    rq_activate_all_grippers(True)
    # end: URCap Program Node
  end
  $ 60 "zero_ftsensor()"
  zero_ftsensor()
  $ 61 "EXTT"
  $ 62 "Set GRP_3F_Enable=Off"
  set_standard_digital_out(4, False)
  $ 63 "Set BarcodeTrigger=Off"
  set_standard_digital_out(6, False)
  $ 64 "Set GRP_3F_Decap=Off"
  set_standard_digital_out(3, False)
  $ 65 "Set GRP_3F_Cap=Off"
  set_standard_digital_out(2, False)
  $ 66 "Set GRP_3F_Open=Off"
  set_standard_digital_out(5, False)
  $ 67 "PSE_T≔get_tool_free_pose(dir=[0,0,0.150], move_in_base_frame=True)"
  global PSE_T=get_tool_free_pose(dir=[0,0,0.150], move_in_base_frame=True)
  $ 68 "If is_reachable(Base_const, [PSE_T])"
  if (is_reachable(p[0.0,0.0,0.0,0.0,0.0,0.0], [PSE_T])):
    $ 69 "MoveL"
    $ 70 "PSE_T" "breakAfter"
    movel(PSE_T, a=1.2, v=0.15)
  end
  $ 71 "powder dispensing variable init"
  $ 72 "Start_thread≔ False "
  global Start_thread=  False
  $ 73 "vib_thread≔ False "
  global vib_thread=  False
  $ 74 "kp≔0.0002"
  global kp=0.0002
  $ 75 "ki≔0.001"
  global ki=0.001
  $ 76 "kd≔0.01"
  global kd=0.01
  $ 77 "dt≔0.05"
  global dt=0.05
  $ 78 "Integral_error≔0"
  global Integral_error=0
  $ 79 "current_error≔0"
  global current_error=0
  $ 80 "previous_error≔0"
  global previous_error=0
  $ 81 "tilt_increment≔0"
  global tilt_increment=0
  $ 82 "tilt_angle≔-1"
  global tilt_angle=-1
  $ 83 "diff≔0"
  global diff=0
  $ 84 "current_pose≔get_actual_tcp_pose()"
  global current_pose= get_actual_tcp_pose ()
  while (True):
    $ 85 "Robot Program"
    $ 86 "MAIN"
    $ 87 "command_manager(external_control='uGO', cond_suspend=(ITM_Manipulated and AMR_AtTarget and AMR_Charging and AMR_Battery<40), cond_unsuspend=(AMR_Battery≟60))"
    command_manager(external_control="uGO", cond_suspend=(ITM_Manipulated  and  AMR_AtTarget  and  AMR_Charging  and  AMR_Battery<40), cond_unsuspend=(AMR_Battery == 60))
    $ 88 "log_state(STATE_Info)"
    log_state(STATE_Info)
    $ 89 "Switch STATE"
    switch_1 = STATE
    $ 90 "Case 1"
    if (1 == switch_1):
      $ 91 "Stopping"
      $ 92 "STATE_Info≔'Stopping'"
      global STATE_Info="Stopping"
      $ 93 "end_freedrive_mode()"
      end_freedrive_mode()
      $ 94 "Set"
      set_tcp(p[0.0,0.0,0.161,3.1415,0.0,0.0])
      $ 95 "PSE_T≔get_tool_free_pose(dir=[0,0,0.150], move_in_base_frame=True)"
      global PSE_T=get_tool_free_pose(dir=[0,0,0.150], move_in_base_frame=True)
      $ 96 "If is_reachable(Base_const, [PSE_T])"
      if (is_reachable(p[0.0,0.0,0.0,0.0,0.0,0.0], [PSE_T])):
        $ 97 "MoveL"
        $ 98 "PSE_T" "breakAfter"
        movel(PSE_T, a=1.2, v=0.15)
      end
      $ 99 "do_transition(keep_rxry=OBJ_Picked, r=0)"
      do_transition(keep_rxry=OBJ_Picked, r=0)
      $ 108 "Call Sub_AMR_MiR_V3"
      Sub_AMR_MiR_V3()
      $ 109 "If stopping() and AMR_Done"
      if (stopping()  and  AMR_Done):
        $ 110 "STATE≔2"
        global STATE=2
        $ 111 "ugo_update_outputs()"
        ugo_update_outputs()
      end
    elif (2 == switch_1):
      $ 112 "Case 2"
      $ 113 "Stopped"
      $ 114 "STATE_Info≔'Stopped'"
      global STATE_Info="Stopped"
      $ 115 "Call Sub_AMR_MiR_V3"
      Sub_AMR_MiR_V3()
      $ 116 "If CMD_Reset  or PB_Start"
      if (CMD_Reset   or  get_standard_digital_in(0)):
        $ 117 "STATE≔3"
        global STATE=3
        $ 118 "ugo_update_outputs()"
        ugo_update_outputs()
      end
    elif (3 == switch_1):
      $ 119 "Case 3"
      $ 120 " Resetting"
      $ 121 "STATE_Info≔'Resetting'"
      global STATE_Info="Resetting"
      $ 122 "uML"
      $ 123 "reset_error()"
      reset_error()
      $ 124 "reset_warning()"
      reset_warning()
      $ 125 "PROCESS_Step≔0"
      global PROCESS_Step=0
      $ 126 "PROCESS_Info≔''"
      global PROCESS_Info=""
      $ 127 "ARM_Referenced≔ False "
      global ARM_Referenced=  False
      $ 128 "WRK_Done≔ False "
      global WRK_Done=  False
      $ 129 "ITM_Prepared≔ False "
      global ITM_Prepared=  False
      $ 130 "ITM_Manipulated≔ False "
      global ITM_Manipulated=  False
      $ 131 "STP≔0"
      global STP=0
      $ 132 "Action≔0"
      global Action=0
      $ 133 "Action_Info≔''"
      global Action_Info=""
      $ 134 "ITM_ID≔0"
      global ITM_ID=0
      $ 135 "JIG≔0"
      global JIG=0
      $ 136 "JIG_Slot≔0"
      global JIG_Slot=0
      $ 137 "Task_info≔''"
      global Task_info=""
      $ 138 "Set"
      set_tcp(p[0.0,0.0,0.161,3.1415,0.0,0.0])
      $ 139 "App"
      $ 140 "'ADD APPLICATION SPECIFIC COMMANDS'"
      # 'ADD APPLICATION SPECIFIC COMMANDS'
      $ 141 "OBJ_Type≔0"
      global OBJ_Type=0
      $ 142 "OBJ_Nbr≔0"
      global OBJ_Nbr=0
      $ 143 "If CNT_Rack_Output≥50"
      if (CNT_Rack_Output >= 50):
        $ 144 "CNT_Rack_Output≔0"
        global CNT_Rack_Output=0
      end
      $ 145 "TASK≔struct(ID=0, NAVI=struct(target=0, footprint=0, protectiveOff=0, dock=0), WORK=struct(ITM_ID_Src=0, JIG_ID_Src=0, OBJ_Nbr_Src=0, ACT_Src=0, ITM_ID_Tgt=0, JIG_ID_Tgt=0, OBJ_Nbr_Tgt=0, ACT_Tgt=0, OBJ_Type=0))"
      global TASK=struct(ID=0, NAVI=struct(target=0, footprint=0, protectiveOff=0, dock=0), WORK=struct(ITM_ID_Src=0, JIG_ID_Src=0, OBJ_Nbr_Src=0, ACT_Src=0, ITM_ID_Tgt=0, JIG_ID_Tgt=0, OBJ_Nbr_Tgt=0, ACT_Tgt=0, OBJ_Type=0))
      $ 146 "Call Sub_AMR_MiR_V3"
      Sub_AMR_MiR_V3()
      $ 147 "If resetting() and AMR_Done"
      if (resetting()  and  AMR_Done):
        $ 148 "STATE≔4"
        global STATE=4
        $ 149 "ugo_update_outputs()"
        ugo_update_outputs()
      end
    elif (4 == switch_1):
      $ 150 "Case 4"
      $ 151 "Idle"
      $ 152 "STATE_Info≔'Idle'"
      global STATE_Info="Idle"
      $ 153 "If CMD_Start"
      if (CMD_Start):
        $ 154 "STATE≔5"
        global STATE=5
        $ 155 "ugo_update_outputs()"
        ugo_update_outputs()
      end
    elif (5 == switch_1):
      $ 156 "Case 5"
      $ 157 "Starting"
      $ 158 "STATE_Info≔'Starting'"
      global STATE_Info="Starting"
      $ 159 "'ADD COMMANDS WHAT TO START WITH'"
      # 'ADD COMMANDS WHAT TO START WITH'
      $ 160 "Call Sub_AMR_MiR_V3"
      Sub_AMR_MiR_V3()
      $ 161 "get ugo data"
      $ 162 "Assign Tasks"
      $ 163 "TASK.ID = ugo_get_task()"
      TASK.ID = ugo_get_task()
      $ 164 "If TASK.ID≟1"
      if (TASK.ID == 1):
        $ 165 "Task_info≔'Charge'"
        global Task_info="Charge"
        $ 166 "Parameters"
        $ 167 "AMR_PosTarget≔1"
        global AMR_PosTarget=1
      else:
        $ 168 "ElseIf TASK.ID≟9"
        if (TASK.ID == 9):
          $ 169 "'Pick Sarstedt Rack from Variable source'"
          # 'Pick Sarstedt Rack from Variable source'
          $ 170 "Task_info≔'Navigate to Target'"
          global Task_info="Navigate to Target"
          $ 171 "Parameters"
          $ 172 "AMR_PosTarget≔UGO.read_input('00','ITM_ID')"
          global AMR_PosTarget=UGO.read_input("00","ITM_ID")
        else:
          $ 173 "ElseIf TASK.ID≟10"
          if (TASK.ID == 10):
            $ 174 "'Pick Sarstedt Rack from Variable source'"
            # 'Pick Sarstedt Rack from Variable source'
            $ 175 "Task_info≔'Pick Rack'"
            global Task_info="Pick Rack"
            $ 176 "AMR_PosTarget≔2"
            global AMR_PosTarget=2
            $ 177 "Parameters"
            $ 178 "ITM_ID≔UGO.read_input('00','ITM_ID')"
            global ITM_ID=UGO.read_input("00","ITM_ID")
            $ 179 "JIG≔UGO.read_input('00','JIG_ID')"
            global JIG=UGO.read_input("00","JIG_ID")
            $ 180 "OBJ_Type≔3"
            global OBJ_Type=3
          else:
            $ 181 "ElseIf TASK.ID≟11"
            if (TASK.ID == 11):
              $ 182 "'Place Sarstedt Rack on Variable target'"
              # 'Place Sarstedt Rack on Variable target'
              $ 183 "Task_info≔'Place Rack'"
              global Task_info="Place Rack"
              $ 184 "AMR_PosTarget≔2"
              global AMR_PosTarget=2
              $ 185 "Parameters"
              $ 186 "ITM_ID≔UGO.read_input('00','ITM_ID')"
              global ITM_ID=UGO.read_input("00","ITM_ID")
              $ 187 "JIG≔UGO.read_input('00','JIG_ID')"
              global JIG=UGO.read_input("00","JIG_ID")
              $ 188 "OBJ_Type≔3"
              global OBJ_Type=3
            else:
              $ 190 "ElseIf TASK.ID≟12"
              if (TASK.ID == 12):
                $ 191 "Task_info≔'Decapping'"
                global Task_info="Decapping"
                $ 192 "Parameters"
                $ 193 "ITM_ID≔1"
                global ITM_ID=1
                $ 194 "AMR_PosTarget≔AMR_PosActual"
                global AMR_PosTarget=AMR_PosActual
                $ 195 "PRC_TubCounter≔0"
                global PRC_TubCounter=0
              else:
                $ 196 "ElseIf TASK.ID≟13"
                if (TASK.ID == 13):
                  $ 197 "Task_info≔'Empty racks'"
                  global Task_info="Empty racks"
                  $ 198 "Parameters"
                  $ 199 "ITM_ID≔1"
                  global ITM_ID=1
                  $ 200 "AMR_PosTarget≔AMR_PosActual"
                  global AMR_PosTarget=AMR_PosActual
                else:
                  $ 201 "ElseIf TASK.ID≟16"
                  if (TASK.ID == 16):
                    $ 202 "Task_info≔'Decap + Barcode'"
                    global Task_info="Decap + Barcode"
                    $ 203 "Parameters"
                    $ 205 "OBJs_String≔UGO.read_input('00','ObjPos')"
                    global OBJs_String=UGO.read_input("00","ObjPos")
                    $ 206 "OBJs_List≔make_list(length = elements_in_string(OBJs_String), initial_value = -1, capacity = 50)"
                    global OBJs_List=make_list(length = elements_in_string(OBJs_String), initial_value = -1, capacity = 50)
                    $ 207 "OBJs_List≔string_to_list(OBJs_String)"
                    global OBJs_List=string_to_list(OBJs_String)
                    $ 208 "ITM_ID≔1"
                    global ITM_ID=1
                    $ 209 "OBJ_Type≔2"
                    global OBJ_Type=2
                    $ 210 "JIG≔7"
                    global JIG=7
                    $ 211 "AMR_PosTarget≔AMR_PosActual"
                    global AMR_PosTarget=AMR_PosActual
                  else:
                    $ 212 "ElseIf TASK.ID≟30"
                    if (TASK.ID == 30):
                      $ 213 "Task_info≔'Getting bottles'"
                      global Task_info="Getting bottles"
                      $ 214 "Parameters"
                      $ 215 "ITM_ID≔1"
                      global ITM_ID=1
                      $ 216 "OBJ_Type≔4"
                      global OBJ_Type=4
                      $ 217 "JIG≔9"
                      global JIG=9
                      $ 218 "AMR_PosTarget≔4"
                      global AMR_PosTarget=4
                    else:
                      $ 219 "ElseIf TASK.ID≟40"
                      if (TASK.ID == 40):
                        $ 220 "Task_info≔'Placing bottles'"
                        global Task_info="Placing bottles"
                        $ 221 "Parameters"
                        $ 222 "ITM_ID≔1"
                        global ITM_ID=1
                        $ 223 "OBJ_Type≔4"
                        global OBJ_Type=4
                        $ 224 "JIG≔10"
                        global JIG=10
                        $ 225 "AMR_PosTarget≔4"
                        global AMR_PosTarget=4
                      else:
                        $ 226 "ElseIf TASK.ID≟41"
                        if (TASK.ID == 41):
                          $ 227 "Task_info≔'Shaking bottle'"
                          global Task_info="Shaking bottle"
                          $ 228 "Parameters"
                          $ 229 "ITM_ID≔1"
                          global ITM_ID=1
                          $ 230 "OBJ_Type≔4"
                          global OBJ_Type=4
                          $ 231 "JIG≔11"
                          global JIG=11
                          $ 232 "AMR_PosTarget≔4"
                          global AMR_PosTarget=4
                        else:
                          $ 233 "ElseIf TASK.ID≟42"
                          if (TASK.ID == 42):
                            $ 234 "Task_info≔'Decap the bottle'"
                            global Task_info="Decap the bottle"
                            $ 235 "Parameters"
                            $ 236 "ITM_ID≔1"
                            global ITM_ID=1
                            $ 237 "OBJ_Type≔4"
                            global OBJ_Type=4
                            $ 238 "AMR_PosTarget≔4"
                            global AMR_PosTarget=4
                          else:
                            $ 239 "ElseIf TASK.ID≟43"
                            if (TASK.ID == 43):
                              $ 240 "Task_info≔'Pick the Rack'"
                              global Task_info="Pick the Rack"
                              $ 241 "AMR_PosTarget≔5"
                              global AMR_PosTarget=5
                              $ 242 "Parameters"
                              $ 243 "ITM_ID≔UGO.read_input('00','ITM_ID')"
                              global ITM_ID=UGO.read_input("00","ITM_ID")
                              $ 244 "JIG≔UGO.read_input('00','JIG_ID')"
                              global JIG=UGO.read_input("00","JIG_ID")
                              $ 245 "OBJ_Type≔3"
                              global OBJ_Type=3
                            else:
                              $ 246 "ElseIf TASK.ID≟45"
                              if (TASK.ID == 45):
                                $ 247 "Task_info≔'pick the Vial'"
                                global Task_info="pick the Vial"
                                $ 248 "Parameters"
                                $ 249 "ITM_ID≔1"
                                global ITM_ID=1
                                $ 250 "OBJ_Type≔4"
                                global OBJ_Type=4
                                $ 251 "JIG≔12"
                                global JIG=12
                                $ 252 "AMR_PosTarget≔5"
                                global AMR_PosTarget=5
                              else:
                                $ 253 "ElseIf TASK.ID≟46"
                                if (TASK.ID == 46):
                                  $ 254 "Task_info≔'Decap the Vial'"
                                  global Task_info="Decap the Vial"
                                  $ 255 "Parameters"
                                  $ 256 "ITM_ID≔1"
                                  global ITM_ID=1
                                  $ 257 "OBJ_Type≔4"
                                  global OBJ_Type=4
                                  $ 258 "JIG≔13"
                                  global JIG=13
                                  $ 259 "AMR_PosTarget≔5"
                                  global AMR_PosTarget=5
                                else:
                                  $ 260 "ElseIf TASK.ID≟47"
                                  if (TASK.ID == 47):
                                    $ 261 "Task_info≔'Liquid Transfer'"
                                    global Task_info="Liquid Transfer"
                                    $ 262 "Parameters"
                                    $ 263 "ITM_ID≔1"
                                    global ITM_ID=1
                                    $ 264 "OBJ_Type≔4"
                                    global OBJ_Type=4
                                    $ 265 "JIG≔14"
                                    global JIG=14
                                    $ 266 "AMR_PosTarget≔3"
                                    global AMR_PosTarget=3
                                  else:
                                    $ 267 "ElseIf TASK.ID≟48"
                                    if (TASK.ID == 48):
                                      $ 268 "Task_info≔'Place_rack'"
                                      global Task_info="Place_rack"
                                      $ 269 "Parameters"
                                      $ 270 "ITM_ID≔1"
                                      global ITM_ID=1
                                      $ 271 "OBJ_Type≔3"
                                      global OBJ_Type=3
                                      $ 272 "JIG≔7"
                                      global JIG=7
                                      $ 273 "AMR_PosTarget≔5"
                                      global AMR_PosTarget=5
                                    else:
                                      $ 274 "ElseIf TASK.ID≟49"
                                      if (TASK.ID == 49):
                                        $ 275 "Task_info≔'Pick Containers'"
                                        global Task_info="Pick Containers"
                                        $ 276 "Parameters"
                                        $ 277 "ITM_ID≔1"
                                        global ITM_ID=1
                                        $ 278 "OBJ_Type≔6"
                                        global OBJ_Type=6
                                        $ 279 "JIG≔15"
                                        global JIG=15
                                        $ 280 "AMR_PosTarget≔3"
                                        global AMR_PosTarget=3
                                      else:
                                        $ 281 "ElseIf TASK.ID≟50"
                                        if (TASK.ID == 50):
                                          $ 282 "Task_info≔'Decap Containers'"
                                          global Task_info="Decap Containers"
                                          $ 283 "Parameters"
                                          $ 284 "ITM_ID≔1"
                                          global ITM_ID=1
                                          $ 285 "OBJ_Type≔6"
                                          global OBJ_Type=6
                                          $ 286 "JIG≔16"
                                          global JIG=16
                                          $ 287 "AMR_PosTarget≔5"
                                          global AMR_PosTarget=5
                                        else:
                                          $ 288 "ElseIf TASK.ID≟51"
                                          if (TASK.ID == 51):
                                            $ 289 "Task_info≔'Detect Spatula and transfer powder'"
                                            global Task_info="Detect Spatula and transfer powder"
                                            $ 290 "Parameters"
                                            $ 291 "ITM_ID≔1"
                                            global ITM_ID=1
                                            $ 292 "OBJ_Type≔8"
                                            global OBJ_Type=8
                                            $ 293 "JIG≔16"
                                            global JIG=16
                                            $ 294 "AMR_PosTarget≔5"
                                            global AMR_PosTarget=5
                                          else:
                                            $ 295 "ElseIf TASK.ID≟99"
                                            if (TASK.ID == 99):
                                              $ 296 "Task_info≔'Decapping and barcode alignment'"
                                              global Task_info="Decapping and barcode alignment"
                                              $ 297 "Parameters"
                                              $ 298 "PRC_TubNumber≔UGO.read_input('00','TubesNb')"
                                              global PRC_TubNumber=UGO.read_input("00","TubesNb")
                                              $ 299 "PRC_TubCounter≔0"
                                              global PRC_TubCounter=0
                                              $ 300 "ITM_ID≔1"
                                              global ITM_ID=1
                                              $ 301 "AMR_PosTarget≔AMR_PosActual"
                                              global AMR_PosTarget=AMR_PosActual
                                            else:
                                              $ 336 "Else" "noBreak"
                                              $ 337 "set_error(ERROR_WRONG_ORDER)"
                                              set_error(ERROR_WRONG_ORDER)
                                            end
                                          end
                                        end
                                      end
                                    end
                                  end
                                end
                              end
                            end
                          end
                        end
                      end
                    end
                  end
                end
              end
            end
          end
        end
      end
      $ 338 "test ugo"
      $ 339 "Wait: 0.2"
      sleep(0.2)
      $ 340 "ugo_update_outputs()"
      ugo_update_outputs()
      $ 341 "If starting() and AMR_Done"
      if (starting()  and  AMR_Done):
        $ 342 "log_message(Task_info, 'New Task: ')"
        log_message(Task_info, "New Task: ")
        $ 343 "log_message(to_str(TASK.ID), 'Task_ID: ')"
        log_message(to_str(TASK.ID), "Task_ID: ")
        $ 344 "do_transition(keep_rxry=OBJ_Picked)"
        do_transition(keep_rxry=OBJ_Picked)
        $ 345 "STATE≔6"
        global STATE=6
        $ 346 "ugo_update_outputs()"
        ugo_update_outputs()
      end
    elif (6 == switch_1):
      $ 347 "Case 6"
      $ 348 "Execute"
      $ 349 "STATE_Info≔'Execute'"
      global STATE_Info="Execute"
      $ 350 "If  not CMD_Hold and not CMD_Suspend"
      global thread_flag_350=0
      thread Thread_if_350():
        $ 351 "Switch PROCESS_Step"
        switch_2 = PROCESS_Step
        $ 352 "Case 0"
        if (0 == switch_2):
          $ 353 "PROCESS_Info≔'process control'"
          global PROCESS_Info="process control"
          $ 354 "log_process(PROCESS_Info)"
          log_process(PROCESS_Info)
          $ 355 "process control"
          $ 356 "If  not AMR_AtTarget"
          if (  not  AMR_AtTarget):
            $ 357 "PROCESS_Step≔1"
            global PROCESS_Step=1
          else:
            $ 358 "ElseIf (( not ITM_Prepared and  not WRK_Done) or (ITM_Prepared and WRK_Done))"
            if (((  not  ITM_Prepared  and    not  WRK_Done)  or  (ITM_Prepared  and  WRK_Done))):
              $ 359 "PROCESS_Step≔2"
              global PROCESS_Step=2
            else:
              $ 360 "ElseIf  not WRK_Done"
              if (  not  WRK_Done):
                $ 361 "PROCESS_Step≔3"
                global PROCESS_Step=3
              else:
                $ 362 "Else" "noBreak"
                $ 363 "task finished"
                $ 364 "PROCESS_Info≔''"
                global PROCESS_Info=""
                $ 365 "STATE≔7"
                global STATE=7
                $ 366 "ugo_update_outputs()"
                ugo_update_outputs()
              end
            end
          end
        elif (1 == switch_2):
          $ 367 "Case 1"
          $ 368 "navigate"
          $ 369 "'MOVING THE uML'"
          # 'MOVING THE uML'
          $ 370 "PROCESS_Info≔'move to target'"
          global PROCESS_Info="move to target"
          $ 371 "log_process(PROCESS_Info)"
          log_process(PROCESS_Info)
          $ 372 "If TASK.ID≟1"
          if (TASK.ID == 1):
            $ 373 "Action≔51"
            global Action=51
          else:
            $ 374 "Else" "noBreak"
            $ 375 "Action≔52"
            global Action=52
          end
          $ 376 "Call Sub_AMR_MiR_V3"
          Sub_AMR_MiR_V3()
          $ 377 "If AMR_Done"
          if (AMR_Done):
            $ 378 "PROCESS_Step≔0"
            global PROCESS_Step=0
          end
        elif (2 == switch_2):
          $ 379 "Case 2"
          $ 380 "prepare"
          $ 381 "'THINGS THAT HAVE TO BE DONE ONCE IN A SEQUENCE,WORKFLOW'"
          # 'THINGS THAT HAVE TO BE DONE ONCE IN A SEQUENCE,WORKFLOW'
          $ 382 "PROCESS_Info≔'prepare for work'"
          global PROCESS_Info="prepare for work"
          $ 383 "log_process(PROCESS_Info)"
          log_process(PROCESS_Info)
          $ 384 "If TASK.WORK.ITM_ID_Src>1"
          if (TASK.WORK.ITM_ID_Src>1):
            $ 385 "ITM_ID≔TASK.WORK.ITM_ID_Src"
            global ITM_ID=TASK.WORK.ITM_ID_Src
          else:
            $ 386 "ElseIf TASK.WORK.ITM_ID_Tgt>1"
            if (TASK.WORK.ITM_ID_Tgt>1):
              $ 387 "ITM_ID≔TASK.WORK.ITM_ID_Tgt"
              global ITM_ID=TASK.WORK.ITM_ID_Tgt
            end
          end
          $ 388 "If  not ARM_Referenced and (ITM_ID≠0)"
          if (  not  ARM_Referenced  and  (ITM_ID != 0)):
            $ 389 "STP≔1"
            global STP=1
          else:
            $ 390 "ElseIf ARM_Referenced or (ITM_ID≟0)"
            if (ARM_Referenced  or  (ITM_ID == 0)):
              $ 391 "STP≔2"
              global STP=2
            end
          end
          $ 392 "Switch STP"
          switch_3 = STP
          $ 393 "Case 1"
          if (1 == switch_3):
            $ 394 "reference"
            $ 395 "STP_Info≔'reference at target position'"
            global STP_Info="reference at target position"
            $ 396 "log_step(STP_Info)"
            log_step(STP_Info)
            $ 397 "If ITM_ID≟1"
            if (ITM_ID == 1):
              $ 398 "CAM_Done≔ True "
              global CAM_Done=  True
            else:
              $ 399 "Else" "noBreak"
              $ 400 "Action≔131"
              global Action=131
              $ 401 "Call Sub_Vision_V18"
              Sub_Vision_V18()
            end
            $ 403 "If CAM_Done and  not ERROR.FLAG"
            if (CAM_Done  and    not  ERROR.FLAG):
              $ 404 "log_step('ARM referenced')"
              log_step("ARM referenced")
              $ 405 "ARM_Referenced≔ True "
              global ARM_Referenced=  True
            end
          elif (2 == switch_3):
            $ 406 "Case 2"
            $ 407 "manipulate"
            $ 408 "STP_Info≔'manipulate item'"
            global STP_Info="manipulate item"
            $ 409 "log_step(STP_Info)"
            log_step(STP_Info)
            $ 410 "'In case pressing button is needed'"
            # 'In case pressing button is needed'
            $ 411 "If found_in_list(ITM_ID, ITM_ID_List)"
            if (found_in_list(ITM_ID, ITM_ID_List)):
              $ 412 "Switch ITM_ID"
              switch_4 = ITM_ID
              $ 413 "Case 0"
              if (0 == switch_4):
                $ 414 "ITM_Manipulated≔ not ITM_Manipulated"
                global ITM_Manipulated=  not  ITM_Manipulated
              elif (1 == switch_4):
                $ 415 "Case 1"
                $ 416 "ITM_Manipulated≔ not ITM_Manipulated"
                global ITM_Manipulated=  not  ITM_Manipulated
              elif (2 == switch_4):
                $ 417 "Case 2"
              else:
                $ 427 "Default Case"
                $ 428 "ITM_Manipulated≔ not ITM_Manipulated"
                global ITM_Manipulated=  not  ITM_Manipulated
              end
            end
          end
          $ 429 "ITM_Prepared≔(ITM_Manipulated or  not found_in_list(ITM_ID, ITM_ID_List)) and (ARM_Referenced or ITM_ID≟0) and  not WRK_Done"
          global ITM_Prepared=(ITM_Manipulated  or    not  found_in_list(ITM_ID, ITM_ID_List))  and  (ARM_Referenced  or  ITM_ID == 0)  and    not  WRK_Done
          $ 430 "STP≔0"
          global STP=0
          $ 431 "STP_Info≔''"
          global STP_Info=""
          $ 432 "PROCESS_Step≔0"
          global PROCESS_Step=0
        elif (3 == switch_2):
          $ 433 "Case 3"
          $ 434 "work"
          $ 435 "'ADD EVERY MACHINE, OBJECT, STATION TO WORK ON'"
          # 'ADD EVERY MACHINE, OBJECT, STATION TO WORK ON'
          $ 436 "Switch ITM_ID"
          switch_3 = ITM_ID
          $ 437 "Case 1"
          if (1 == switch_3):
            $ 438 "uLM"
            $ 439 "If TASK.ID≟12"
            if (TASK.ID == 12):
              $ 440 "fill racks"
              $ 441 "Action≔151"
              global Action=151
              $ 442 "Call Sub_Vision_V18"
              Sub_Vision_V18()
              $ 443 "If  not ERROR.FLAG"
              if (  not  ERROR.FLAG):
                $ 444 "Actions for the task"
                $ 445 "Action≔1"
                global Action=1
                $ 446 "JIG≔2"
                global JIG=2
                $ 447 "JIG_Slot≔CAM_Result[0]"
                global JIG_Slot=CAM_Result[0]
                $ 448 "OBJ_Nbr≔CAM_Result[0]"
                global OBJ_Nbr=CAM_Result[0]
                $ 449 "OBJ_Type≔2"
                global OBJ_Type=2
                $ 450 "Call Sub_Action_V4"
                Sub_Action_V4()
                $ 451 "If OBJ_Picked"
                if (OBJ_Picked):
                  $ 452 "CAM_Result.remove(0)"
                  CAM_Result.remove(0)
                  $ 453 "PRC_TubCounter≔PRC_TubCounter+1"
                  global PRC_TubCounter=PRC_TubCounter+1
                  $ 454 "If PRC_TubCounter%4≟0"
                  if (PRC_TubCounter%4 == 0):
                    $ 455 "JIG_Slot≔4"
                    global JIG_Slot=4
                  else:
                    $ 456 "Else" "noBreak"
                    $ 457 "JIG_Slot≔PRC_TubCounter%4"
                    global JIG_Slot=PRC_TubCounter%4
                  end
                  $ 458 "OBJ_Nbr≔ceil(PRC_TubCounter/4)"
                  global OBJ_Nbr=ceil(PRC_TubCounter/4)
                  $ 459 "Action≔2"
                  global Action=2
                  $ 460 "JIG≔4"
                  global JIG=4
                  $ 461 "Call Sub_Action_V4"
                  Sub_Action_V4()
                  $ 462 "Action≔151"
                  global Action=151
                  $ 463 "Call Sub_Vision_V18"
                  Sub_Vision_V18()
                end
              end
              $ 464 "If (CAM_Captures≥CAM_PRM_Retries) or (PRC_TubCounter≥32)"
              if ((CAM_Captures >= CAM_PRM_Retries)  or  (PRC_TubCounter >= 32)):
                $ 465 "PROCESS_Step≔0"
                global PROCESS_Step=0
                $ 466 "WRK_Done≔ True "
                global WRK_Done=  True
              end
            else:
              $ 467 "ElseIf TASK.ID≟10"
              if (TASK.ID == 10):
                $ 468 "Pick Rack"
                $ 469 "Action≔131"
                global Action=131
                $ 470 "Call Sub_Vision_V18"
                Sub_Vision_V18()
                $ 471 "Action≔1"
                global Action=1
                $ 472 "Call Sub_Action_V4"
                Sub_Action_V4()
                $ 473 "PROCESS_Step≔0"
                global PROCESS_Step=0
                $ 474 "WRK_Done≔ True "
                global WRK_Done=  True
              else:
                $ 475 "ElseIf TASK.ID≟11"
                if (TASK.ID == 11):
                  $ 476 "Place Rack"
                  $ 477 "Action≔2"
                  global Action=2
                  $ 478 "Call Sub_Action_V4"
                  Sub_Action_V4()
                  $ 479 "PROCESS_Step≔0"
                  global PROCESS_Step=0
                  $ 480 "WRK_Done≔ True "
                  global WRK_Done=  True
                else:
                  $ 481 "ElseIf TASK.ID≟13"
                  if (TASK.ID == 13):
                    $ 482 "empty racks"
                    $ 483 "pick"
                    $ 484 "Action≔1"
                    global Action=1
                    $ 485 "JIG≔4"
                    global JIG=4
                    $ 486 "If PRC_TubCounter%4≟0"
                    if (PRC_TubCounter%4 == 0):
                      $ 487 "JIG_Slot≔4"
                      global JIG_Slot=4
                    else:
                      $ 488 "Else" "noBreak"
                      $ 489 "JIG_Slot≔PRC_TubCounter%4"
                      global JIG_Slot=PRC_TubCounter%4
                    end
                    $ 490 "OBJ_Nbr≔ceil(PRC_TubCounter/4)"
                    global OBJ_Nbr=ceil(PRC_TubCounter/4)
                    $ 491 "OBJ_Type≔2"
                    global OBJ_Type=2
                    $ 492 "Call Sub_Action_V4"
                    Sub_Action_V4()
                    $ 493 "If OBJ_Picked"
                    if (OBJ_Picked):
                      $ 494 "Action≔2"
                      global Action=2
                      $ 495 "JIG≔3"
                      global JIG=3
                      $ 496 "JIG_Slot≔1"
                      global JIG_Slot=1
                      $ 497 "CNT_Rack_Output≔CNT_Rack_Output + 1"
                      global CNT_Rack_Output=CNT_Rack_Output + 1
                      $ 498 "OBJ_Nbr≔CNT_Rack_Output"
                      global OBJ_Nbr=CNT_Rack_Output
                      $ 499 "Call Sub_Action_V4"
                      Sub_Action_V4()
                      $ 500 "If  not ERROR.FLAG"
                      if (  not  ERROR.FLAG):
                        $ 501 "PRC_TubCounter≔PRC_TubCounter - 1"
                        global PRC_TubCounter=PRC_TubCounter - 1
                      end
                    end
                    $ 502 "If CNT_Rack_Output≥50 or PRC_TubCounter≤0"
                    if (CNT_Rack_Output >= 50  or  PRC_TubCounter <= 0):
                      $ 503 "PROCESS_Step≔0"
                      global PROCESS_Step=0
                      $ 504 "WRK_Done≔ True "
                      global WRK_Done=  True
                    end
                  else:
                    $ 505 "ElseIf TASK.ID≟16"
                    if (TASK.ID == 16):
                      $ 506 "CAM_Result≔OBJs_List"
                      global CAM_Result=OBJs_List
                      $ 507 "PRC_CntDetect≔0"
                      global PRC_CntDetect=0
                      $ 508 "Loop PRC_CntDetect<CAM_Result.length()"
                      while (PRC_CntDetect<CAM_Result.length()):
                        $ 509 "Action≔1"
                        global Action=1
                        $ 510 "ITM_ID≔1"
                        global ITM_ID=1
                        $ 511 "JIG≔2"
                        global JIG=2
                        $ 512 "OBJ_Type≔2"
                        global OBJ_Type=2
                        $ 513 "JIG_Slot≔CAM_Result[PRC_CntDetect]"
                        global JIG_Slot=CAM_Result[PRC_CntDetect]
                        $ 514 "OBJ_Nbr≔CAM_Result[PRC_CntDetect]"
                        global OBJ_Nbr=CAM_Result[PRC_CntDetect]
                        $ 515 "Call Sub_Action_V4"
                        Sub_Action_V4()
                        $ 516 "JIG≔1"
                        global JIG=1
                        $ 517 "Action≔11"
                        global Action=11
                        $ 518 "Call Sub_Action_V4"
                        Sub_Action_V4()
                        $ 519 "Action≔12"
                        global Action=12
                        $ 520 "Call Sub_Action_V4"
                        Sub_Action_V4()
                        $ 521 "Action≔6"
                        global Action=6
                        $ 522 "JIG≔6"
                        global JIG=6
                        $ 523 "Call Sub_Action_V4"
                        Sub_Action_V4()
                        $ 524 "Action≔13"
                        global Action=13
                        $ 525 "Call Sub_Action_V4"
                        Sub_Action_V4()
                        $ 526 "Action≔1"
                        global Action=1
                        $ 527 "JIG≔1"
                        global JIG=1
                        $ 528 "Call Sub_Action_V4"
                        Sub_Action_V4()
                        $ 529 "If OBJ_Brc_OK"
                        if (OBJ_Brc_OK):
                          $ 530 "JIG≔2"
                          global JIG=2
                          $ 531 "Action≔2"
                          global Action=2
                          $ 532 "OBJ_Nbr≔CAM_Result[PRC_CntDetect]"
                          global OBJ_Nbr=CAM_Result[PRC_CntDetect]
                          $ 533 "JIG_Slot≔CAM_Result[PRC_CntDetect]"
                          global JIG_Slot=CAM_Result[PRC_CntDetect]
                          $ 534 "OBJ_Type≔2"
                          global OBJ_Type=2
                          $ 535 "Call Sub_Action_V4"
                          Sub_Action_V4()
                        else:
                          $ 536 "Else" "noBreak"
                          $ 537 "Action≔2"
                          global Action=2
                          $ 538 "JIG≔8"
                          global JIG=8
                          $ 539 "Call Sub_Action_V4"
                          Sub_Action_V4()
                        end
                        $ 540 "PRC_CntDetect≔PRC_CntDetect+1"
                        global PRC_CntDetect=PRC_CntDetect+1
                      end
                      $ 541 "PROCESS_Step≔0"
                      global PROCESS_Step=0
                      $ 542 "WRK_Done≔ True "
                      global WRK_Done=  True
                    else:
                      $ 543 "ElseIf TASK.ID≟30"
                      if (TASK.ID == 30):
                        $ 544 "Pick Bottle"
                        $ 545 "Action≔1"
                        global Action=1
                        $ 546 "Call Sub_Action_V4"
                        Sub_Action_V4()
                        $ 547 "PROCESS_Step≔0"
                        global PROCESS_Step=0
                        $ 548 "WRK_Done≔ True "
                        global WRK_Done=  True
                      else:
                        $ 549 "ElseIf TASK.ID≟40"
                        if (TASK.ID == 40):
                          $ 550 "Place Bottle"
                          $ 551 "Action≔2"
                          global Action=2
                          $ 552 "Call Sub_Action_V4"
                          Sub_Action_V4()
                          $ 553 "PROCESS_Step≔0"
                          global PROCESS_Step=0
                          $ 554 "WRK_Done≔ True "
                          global WRK_Done=  True
                        else:
                          $ 555 "ElseIf TASK.ID≟45"
                          if (TASK.ID == 45):
                            $ 556 "Pick Vial"
                            $ 557 "Action≔31"
                            global Action=31
                            $ 558 "Call Sub_Action_V4"
                            Sub_Action_V4()
                            $ 559 "PROCESS_Step≔0"
                            global PROCESS_Step=0
                            $ 560 "WRK_Done≔ True "
                            global WRK_Done=  True
                          else:
                            $ 561 "ElseIf TASK.ID≟46"
                            if (TASK.ID == 46):
                              $ 562 "Decap Vial"
                              $ 563 "Action≔32"
                              global Action=32
                              $ 564 "Call Sub_Action_V4"
                              Sub_Action_V4()
                              $ 565 "PROCESS_Step≔0"
                              global PROCESS_Step=0
                              $ 566 "WRK_Done≔ True "
                              global WRK_Done=  True
                            else:
                              $ 567 "ElseIf TASK.ID≟47"
                              if (TASK.ID == 47):
                                $ 568 "Liquid transfer"
                                $ 569 "Action≔33"
                                global Action=33
                                $ 570 "Call Sub_Action_V4"
                                Sub_Action_V4()
                                $ 571 "PROCESS_Step≔0"
                                global PROCESS_Step=0
                                $ 572 "WRK_Done≔ True "
                                global WRK_Done=  True
                              else:
                                $ 573 "ElseIf TASK.ID≟48"
                                if (TASK.ID == 48):
                                  $ 574 "Place Rack"
                                  $ 575 "Action≔34"
                                  global Action=34
                                  $ 576 "Call Sub_Action_V4"
                                  Sub_Action_V4()
                                  $ 577 "PROCESS_Step≔0"
                                  global PROCESS_Step=0
                                  $ 578 "WRK_Done≔ True "
                                  global WRK_Done=  True
                                else:
                                  $ 579 "ElseIf TASK.ID≟49"
                                  if (TASK.ID == 49):
                                    $ 580 "Pick Powder container"
                                    $ 581 "Action≔35"
                                    global Action=35
                                    $ 582 "Call Sub_Action_V4"
                                    Sub_Action_V4()
                                    $ 583 "PROCESS_Step≔0"
                                    global PROCESS_Step=0
                                    $ 584 "WRK_Done≔ True "
                                    global WRK_Done=  True
                                  else:
                                    $ 585 "ElseIf TASK.ID≟41"
                                    if (TASK.ID == 41):
                                      $ 586 "shake Bottle"
                                      $ 587 "Action≔30"
                                      global Action=30
                                      $ 588 "Call Sub_Action_V4"
                                      Sub_Action_V4()
                                      $ 589 "PROCESS_Step≔0"
                                      global PROCESS_Step=0
                                      $ 590 "WRK_Done≔ True "
                                      global WRK_Done=  True
                                    else:
                                      $ 591 "ElseIf TASK.ID≟42"
                                      if (TASK.ID == 42):
                                        $ 592 "decap the bottle"
                                        $ 593 "Action≔1"
                                        global Action=1
                                        $ 594 "JIG≔9"
                                        global JIG=9
                                        $ 595 "Call Sub_Action_V4"
                                        Sub_Action_V4()
                                        $ 596 "Action≔11"
                                        global Action=11
                                        $ 597 "JIG≔1"
                                        global JIG=1
                                        $ 598 "Call Sub_Action_V4"
                                        Sub_Action_V4()
                                        $ 599 "Action≔12"
                                        global Action=12
                                        $ 600 "JIG≔1"
                                        global JIG=1
                                        $ 601 "Call Sub_Action_V4"
                                        Sub_Action_V4()
                                        $ 602 "Action≔2"
                                        global Action=2
                                        $ 603 "JIG≔8"
                                        global JIG=8
                                        $ 604 "Call Sub_Action_V4"
                                        Sub_Action_V4()
                                        $ 605 "PROCESS_Step≔0"
                                        global PROCESS_Step=0
                                        $ 606 "WRK_Done≔ True "
                                        global WRK_Done=  True
                                      else:
                                        $ 607 "ElseIf TASK.ID≟43"
                                        if (TASK.ID == 43):
                                          $ 608 "Pick the rack"
                                          $ 609 "Action≔131"
                                          global Action=131
                                          $ 610 "Call Sub_Vision_V18"
                                          Sub_Vision_V18()
                                          $ 611 "Action≔1"
                                          global Action=1
                                          $ 612 "Call Sub_Action_V4"
                                          Sub_Action_V4()
                                          $ 613 "PROCESS_Step≔0"
                                          global PROCESS_Step=0
                                          $ 614 "WRK_Done≔ True "
                                          global WRK_Done=  True
                                        else:
                                          $ 615 "ElseIf TASK.ID≟50"
                                          if (TASK.ID == 50):
                                            $ 616 "Decap containers"
                                            $ 617 "Action≔36"
                                            global Action=36
                                            $ 618 "Call Sub_Action_V4"
                                            Sub_Action_V4()
                                            $ 619 "PROCESS_Step≔0"
                                            global PROCESS_Step=0
                                            $ 620 "WRK_Done≔ True "
                                            global WRK_Done=  True
                                          else:
                                            $ 621 "ElseIf TASK.ID≟51"
                                            if (TASK.ID == 51):
                                              $ 622 "Detect Spatula and transfer powder"
                                              $ 623 "Action≔37"
                                              global Action=37
                                              $ 624 "Call Sub_Action_V4"
                                              Sub_Action_V4()
                                              $ 625 "PROCESS_Step≔0"
                                              global PROCESS_Step=0
                                              $ 626 "WRK_Done≔ True "
                                              global WRK_Done=  True
                                            end
                                          end
                                        end
                                      end
                                    end
                                  end
                                end
                              end
                            end
                          end
                        end
                      end
                    end
                  end
                end
              end
            end
          elif (2 == switch_3):
            $ 627 "Case 2"
          elif (5 == switch_3):
            $ 669 "Case 5"
            $ 670 "SarstedtTable"
            $ 671 "Action≔131"
            global Action=131
            $ 672 "Call Sub_Vision_V18"
            Sub_Vision_V18()
            $ 673 "Action≔1"
            global Action=1
            $ 674 "Call Sub_Action_V4"
            Sub_Action_V4()
            $ 675 "PROCESS_Step≔0"
            global PROCESS_Step=0
            $ 676 "WRK_Done≔ True "
            global WRK_Done=  True
          elif (20 == switch_3):
            $ 677 "Case 20"
          elif (43 == switch_3):
            $ 739 "Case 43"
            $ 740 "Pick the rack"
            $ 741 "Action≔131"
            global Action=131
            $ 742 "Call Sub_Vision_V18"
            Sub_Vision_V18()
            $ 743 "Action≔1"
            global Action=1
            $ 744 "Call Sub_Action_V4"
            Sub_Action_V4()
            $ 745 "PROCESS_Step≔0"
            global PROCESS_Step=0
            $ 746 "WRK_Done≔ True "
            global WRK_Done=  True
          else:
            $ 747 "Default Case"
            $ 748 "WRK_Done≔ True "
            global WRK_Done=  True
            $ 749 "PROCESS_Step≔0"
            global PROCESS_Step=0
          end
        end
        thread_flag_350 = 1
      end
      if (  not  CMD_Hold and not CMD_Suspend):
        global thread_handler_350=run Thread_if_350()
        while (thread_flag_350 == 0):
          if not(  not  CMD_Hold and not CMD_Suspend):
            kill thread_handler_350
            thread_flag_350 = 2
          else:
            sync()
          end
        end
      else:
        thread_flag_350 = 2
      end
      $ 750 "If CMD_Hold"
      if (CMD_Hold):
        $ 751 "STATE≔9"
        global STATE=9
        $ 752 "ugo_update_outputs()"
        ugo_update_outputs()
      else:
        $ 753 "ElseIf CMD_Suspend"
        if (CMD_Suspend):
          $ 754 "STATE≔12"
          global STATE=12
          $ 755 "ugo_update_outputs()"
          ugo_update_outputs()
        end
      end
    elif (7 == switch_1):
      $ 756 "Case 7"
      $ 757 "Completing"
      $ 758 "STATE_Info≔'Completing'"
      global STATE_Info="Completing"
      $ 759 "'ADD COMMANDS FOR COMPLETING THE PROCESS'"
      # 'ADD COMMANDS FOR COMPLETING THE PROCESS'
      $ 760 "do_transition(keep_rxry=OBJ_Picked)"
      do_transition(keep_rxry=OBJ_Picked)
      $ 761 "Call Sub_AMR_MiR_V3"
      Sub_AMR_MiR_V3()
      $ 762 "If completing() and AMR_Done"
      if (completing()  and  AMR_Done):
        $ 763 "STATE≔8"
        global STATE=8
        $ 764 "ugo_update_outputs()"
        ugo_update_outputs()
      end
    elif (8 == switch_1):
      $ 765 "Case 8"
      $ 766 "Complete"
      $ 767 "STATE_Info≔'Complete'"
      global STATE_Info="Complete"
      $ 768 "If CMD_Reset"
      if (CMD_Reset):
        $ 769 "STATE≔3"
        global STATE=3
        $ 770 "ugo_update_outputs()"
        ugo_update_outputs()
      end
    elif (9 == switch_1):
      $ 771 "Case 9"
      $ 772 "Holding"
      $ 773 "STATE_Info≔'Holding'"
      global STATE_Info="Holding"
      $ 774 "stopl(0.5)"
      stopl(0.5)
      $ 775 "Call Sub_AMR_MiR_V3"
      Sub_AMR_MiR_V3()
      $ 776 "If holding() and AMR_Done"
      if (holding()  and  AMR_Done):
        $ 777 "STATE≔10"
        global STATE=10
        $ 778 "ugo_update_outputs()"
        ugo_update_outputs()
      end
    elif (10 == switch_1):
      $ 779 "Case 10"
      $ 780 "Held"
      $ 781 "STATE_Info≔'Held'"
      global STATE_Info="Held"
      $ 782 "If CMD_Unhold"
      if (CMD_Unhold):
        $ 783 "end_freedrive_mode()"
        end_freedrive_mode()
        $ 784 "STATE≔11"
        global STATE=11
        $ 785 "ugo_update_outputs()"
        ugo_update_outputs()
      else:
        $ 786 "ElseIf FNC_Freedrive"
        if (FNC_Freedrive):
          $ 787 "freedrive_mode()"
          freedrive_mode()
        else:
          $ 788 "Else" "noBreak"
          $ 789 "end_freedrive_mode()"
          end_freedrive_mode()
        end
      end
    elif (11 == switch_1):
      $ 790 "Case 11"
      $ 791 "Unholding"
      $ 792 "STATE_Info≔'Unholding'"
      global STATE_Info="Unholding"
      $ 793 "Clearing"
      $ 794 "Switch ERROR.ID"
      switch_2 = ERROR.ID
      $ 795 "Case 1002"
      if (1002 == switch_2):
        $ 796 "AMR_AtTarget≔ False "
        global AMR_AtTarget=  False
        $ 797 "ARM_Referenced≔ False "
        global ARM_Referenced=  False
        $ 798 "ITM_Prepared≔ False "
        global ITM_Prepared=  False
        $ 799 "PROCESS_Step≔1"
        global PROCESS_Step=1
      elif (2007 == switch_2):
        $ 800 "Case 2007"
        $ 801 "PROCESS_Step≔1"
        global PROCESS_Step=1
      end
      $ 802 "reset_error()"
      reset_error()
      $ 803 "reset_warning()"
      reset_warning()
      $ 804 "OBJ_Picked≔gripper_has_object()"
      global OBJ_Picked=gripper_has_object()
      $ 805 "Call Sub_AMR_MiR_V3"
      Sub_AMR_MiR_V3()
      $ 806 "If unholding() and AMR_Done"
      if (unholding()  and  AMR_Done):
        $ 807 "STATE≔6"
        global STATE=6
        $ 808 "ugo_update_outputs()"
        ugo_update_outputs()
      end
    elif (12 == switch_1):
      $ 809 "Case 12"
      $ 810 "Suspending"
      $ 811 "STATE_Info≔'Suspending'"
      global STATE_Info="Suspending"
      $ 812 "PROCESS_Info≔str_cat(PROCESS_Info, ' suspended')"
      global PROCESS_Info=str_cat(PROCESS_Info, " suspended")
      $ 813 "If suspending()"
      if (suspending()):
        $ 814 "STATE≔13"
        global STATE=13
        $ 815 "ugo_update_outputs()"
        ugo_update_outputs()
      end
    elif (13 == switch_1):
      $ 816 "Case 13"
      $ 817 "Suspended"
      $ 818 "STATE_Info≔'Suspended'"
      global STATE_Info="Suspended"
      $ 819 "Call Sub_AMR_MiR_V3"
      Sub_AMR_MiR_V3()
      $ 820 "If CMD_Unsuspend"
      if (CMD_Unsuspend):
        $ 821 "STATE≔14"
        global STATE=14
        $ 822 "ugo_update_outputs()"
        ugo_update_outputs()
      end
    elif (14 == switch_1):
      $ 823 "Case 14"
      $ 824 "Unsuspending"
      $ 825 "STATE_Info≔'Unsuspending'"
      global STATE_Info="Unsuspending"
      $ 826 "PROCESS_Step≔0"
      global PROCESS_Step=0
      $ 827 "If unsuspending()"
      if (unsuspending()):
        $ 828 "STATE≔6"
        global STATE=6
        $ 829 "ugo_update_outputs()"
        ugo_update_outputs()
      end
    elif (15 == switch_1):
      $ 830 "Case 15"
      $ 831 "Aborting"
      $ 832 "STATE_Info≔'Aborting'"
      global STATE_Info="Aborting"
      $ 833 "If aborting()"
      if (aborting()):
        $ 834 "STATE≔16"
        global STATE=16
        $ 835 "ugo_update_outputs()"
        ugo_update_outputs()
      end
    elif (16 == switch_1):
      $ 836 "Case 16"
      $ 837 "Aborted"
      $ 838 "STATE_Info≔'Aborted'"
      global STATE_Info="Aborted"
      $ 839 "If CMD_Clear"
      if (CMD_Clear):
        $ 840 "STATE≔17"
        global STATE=17
        $ 841 "ugo_update_outputs()"
        ugo_update_outputs()
      end
    elif (17 == switch_1):
      $ 842 "Case 17"
      $ 843 "Clearing"
      $ 844 "STATE_Info≔'Clearing'"
      global STATE_Info="Clearing"
      $ 845 "Clearing"
      $ 846 "reset_warning()"
      reset_warning()
      $ 847 "reset_error()"
      reset_error()
      $ 848 "If clearing()"
      if (clearing()):
        $ 849 "STATE≔2"
        global STATE=2
        $ 850 "ugo_update_outputs()"
        ugo_update_outputs()
      end
    end
    $ 851 "log_state(STATE_Info)"
    log_state(STATE_Info)
    $ 852 "log_warning(WARNING.MSG)"
    log_warning(WARNING.MSG)
    $ 853 "log_error(ERROR.MSG)"
    log_error(ERROR.MSG)
    $ 854 "Times"
    $ 855 "Switch STATE"
    switch_1 = STATE
    $ 856 "Case 1"
    if (1 == switch_1):
      $ 857 "TM_St_Stopping≔get_time(STATE_Times[STATE-1])"
      global TM_St_Stopping=get_time(STATE_Times[STATE-1])
    elif (2 == switch_1):
      $ 858 "Case 2"
      $ 859 "TM_St_Stopped≔get_time(STATE_Times[STATE-1])"
      global TM_St_Stopped=get_time(STATE_Times[STATE-1])
    elif (3 == switch_1):
      $ 860 "Case 3"
      $ 861 "TM_St_Resetting≔get_time(STATE_Times[STATE-1])"
      global TM_St_Resetting=get_time(STATE_Times[STATE-1])
    elif (4 == switch_1):
      $ 862 "Case 4"
      $ 863 "TM_St_Idle≔get_time(STATE_Times[STATE-1])"
      global TM_St_Idle=get_time(STATE_Times[STATE-1])
    elif (5 == switch_1):
      $ 864 "Case 5"
      $ 865 "TM_St_Starting≔get_time(STATE_Times[STATE-1])"
      global TM_St_Starting=get_time(STATE_Times[STATE-1])
    elif (6 == switch_1):
      $ 866 "Case 6"
      $ 867 "TM_St_Execute≔get_time(STATE_Times[STATE-1])"
      global TM_St_Execute=get_time(STATE_Times[STATE-1])
    elif (7 == switch_1):
      $ 868 "Case 7"
      $ 869 "TM_St_Completin≔get_time(STATE_Times[STATE-1])"
      global TM_St_Completin=get_time(STATE_Times[STATE-1])
    elif (8 == switch_1):
      $ 870 "Case 8"
      $ 871 "TM_St_Complete≔get_time(STATE_Times[STATE-1])"
      global TM_St_Complete=get_time(STATE_Times[STATE-1])
    elif (9 == switch_1):
      $ 872 "Case 9"
      $ 873 "TM_St_Holding≔get_time(STATE_Times[STATE-1])"
      global TM_St_Holding=get_time(STATE_Times[STATE-1])
    elif (10 == switch_1):
      $ 874 "Case 10"
      $ 875 "TM_St_Held≔get_time(STATE_Times[STATE-1])"
      global TM_St_Held=get_time(STATE_Times[STATE-1])
    elif (11 == switch_1):
      $ 876 "Case 11"
      $ 877 "TM_St_Unholding≔get_time(STATE_Times[STATE-1])"
      global TM_St_Unholding=get_time(STATE_Times[STATE-1])
    elif (12 == switch_1):
      $ 878 "Case 12"
      $ 879 "TM_St_Suspendin≔get_time(STATE_Times[STATE-1])"
      global TM_St_Suspendin=get_time(STATE_Times[STATE-1])
    elif (13 == switch_1):
      $ 880 "Case 13"
      $ 881 "TM_St_Suspended≔get_time(STATE_Times[STATE-1])"
      global TM_St_Suspended=get_time(STATE_Times[STATE-1])
    elif (14 == switch_1):
      $ 882 "Case 14"
      $ 883 "TM_St_Unsuspend≔get_time(STATE_Times[STATE-1])"
      global TM_St_Unsuspend=get_time(STATE_Times[STATE-1])
    elif (15 == switch_1):
      $ 884 "Case 15"
      $ 885 "TM_St_Aborting≔get_time(STATE_Times[STATE-1])"
      global TM_St_Aborting=get_time(STATE_Times[STATE-1])
    elif (16 == switch_1):
      $ 886 "Case 16"
      $ 887 "TM_St_Aborted≔get_time(STATE_Times[STATE-1])"
      global TM_St_Aborted=get_time(STATE_Times[STATE-1])
    elif (17 == switch_1):
      $ 888 "Case 17"
      $ 889 "TM_St_Clearing≔get_time(STATE_Times[STATE-1])"
      global TM_St_Clearing=get_time(STATE_Times[STATE-1])
    end
    $ 891 "Wait: 0.1"
    sleep(0.1)
  end
end
